            "FRK_SetRuntime".Work[#RootIndex].Payload.Info.RecordCount := #Slot;
        ELSIF #Phase = 2 THEN
            #Slot := "FRK_SetRecord"(RootIndex := #RootIndex, Scope := #Status.Name, WriteKey := "FRK_ConfigScratch".Entry.WriteKey);
            #Stored := "FRK_SetRuntime".Work[#RootIndex].Targets[#Slot];
            "FRK_ConfigCommit"(SlotIndex := #Stored, ModelCode := "FRK_SetRuntime".Work[#RootIndex].Payload.Info.ModelCode, Schema := "FRK_ConfigScratch".Schema, Record := "FRK_SetRuntime".Work[#RootIndex].Payload.Records[#Slot]);
        ELSE
            #Slot := "FRK_SetCheck"(RootIndex := #RootIndex, Scope := #Status.Name, Access := #Access, Ready := #Ready, WriteAccess := #Phase <> 3, ReserveTarget := #Phase = 1);
            IF #Slot = 0 THEN RETURN; END_IF;
            IF #Phase = 1 THEN
    #ConfigStageStationCfg.RequireTwoHandStart := "FRK_ConfigScratch".Value.Flag;
            END_IF;
        END_IF;
    END_IF;
    IF "FRK_SetRuntime".Work[#RootIndex].Payload.Info.Kind = 0 THEN
        "FRK_CfgDef_PressDemoUnit"(FieldIndex := 3);
        "FRK_SetRuntime".Work[#RootIndex].RejectScope := #Status.Name;
        "FRK_SetRuntime".Work[#RootIndex].RejectKey := "FRK_ConfigScratch".Entry.WriteKey;
        IF #Phase = 0 OR #Phase = 5 THEN
            IF #Phase = 5 AND NOT "FRK_ConfigDataAllowed"(Access := #Access, ForWrite := FALSE, Scope := #Status.Name) THEN RETURN; END_IF;
            IF #Phase = 5 AND (0 <> 0 OR "FRK_SetRuntime".Work[#RootIndex].Payload.Info.ModelCode = "FRK_ConfigStore".ActiveModels[#RootIndex]) THEN
    "FRK_ConfigScratch".Entry.ValueText := UDINT_TO_WSTRING(#ParCfg.IdealCycleMs);
                #Ok := "FRK_ConfigValidate"(Text := "FRK_ConfigScratch".Entry.ValueText);
            ELSE
                #Ok := "FRK_ConfigGet"(Scope := #Status.Name, ModelCode := "FRK_SetRuntime".Work[#RootIndex].Payload.Info.ModelCode);
            END_IF;
            IF NOT #Ok OR "FRK_SetRuntime".Work[#RootIndex].Payload.Info.RecordCount >= 21 THEN RETURN; END_IF;
            #Slot := "FRK_SetRuntime".Work[#RootIndex].Payload.Info.RecordCount + 1;
            "FRK_SetRuntime".Work[#RootIndex].Payload.Records[#Slot].Scope := #Status.Name;
            "FRK_SetRuntime".Work[#RootIndex].Payload.Records[#Slot].WriteKey := "FRK_ConfigScratch".Entry.WriteKey;
            "FRK_SetRuntime".Work[#RootIndex].Payload.Records[#Slot].Revision := "FRK_ConfigScratch".Entry.WriteRevision;
            "FRK_SetRuntime".Work[#RootIndex].Payload.Records[#Slot].Kind := "FRK_ConfigScratch".Entry.ConfigKind;
            "FRK_SetRuntime".Work[#RootIndex].Payload.Records[#Slot].ValueType := "FRK_ConfigScratch".Entry.ValueType;
            "FRK_SetRuntime".Work[#RootIndex].Payload.Records[#Slot].ValueText := WSTRING_TO_STRING("FRK_ConfigScratch".Entry.ValueText);
            "FRK_SetRuntime".Work[#RootIndex].Payload.Info.RecordCount := #Slot;
        ELSIF #Phase = 2 THEN
            #Slot := "FRK_SetRecord"(RootIndex := #RootIndex, Scope := #Status.Name, WriteKey := "FRK_ConfigScratch".Entry.WriteKey);
            #Stored := "FRK_SetRuntime".Work[#RootIndex].Targets[#Slot];
            "FRK_ConfigCommit"(SlotIndex := #Stored, ModelCode := "FRK_SetRuntime".Work[#RootIndex].Payload.Info.ModelCode, Schema := "FRK_ConfigScratch".Schema, Record := "FRK_SetRuntime".Work[#RootIndex].Payload.Records[#Slot]);
        ELSE
            #Slot := "FRK_SetCheck"(RootIndex := #RootIndex, Scope := #Status.Name, Access := #Access, Ready := #Ready, WriteAccess := #Phase <> 3, ReserveTarget := #Phase = 1);
            IF #Slot = 0 THEN RETURN; END_IF;
            IF #Phase = 1 THEN
    #ConfigStageParCfg.IdealCycleMs := LINT_TO_UDINT("FRK_ConfigScratch".Value.Number);
            END_IF;
        END_IF;
    END_IF;
    IF "FRK_SetRuntime".Work[#RootIndex].Payload.Info.Kind = 0 THEN
        "FRK_CfgDef_PressDemoUnit"(FieldIndex := 4);
        "FRK_SetRuntime".Work[#RootIndex].RejectScope := #Status.Name;
        "FRK_SetRuntime".Work[#RootIndex].RejectKey := "FRK_ConfigScratch".Entry.WriteKey;
        IF #Phase = 0 OR #Phase = 5 THEN
            IF #Phase = 5 AND NOT "FRK_ConfigDataAllowed"(Access := #Access, ForWrite := FALSE, Scope := #Status.Name) THEN RETURN; END_IF;
            IF #Phase = 5 AND (0 <> 0 OR "FRK_SetRuntime".Work[#RootIndex].Payload.Info.ModelCode = "FRK_ConfigStore".ActiveModels[#RootIndex]) THEN
    "FRK_ConfigScratch".Entry.ValueText := UDINT_TO_WSTRING(#ParCfg.BaselineWorkMs);
                #Ok := "FRK_ConfigValidate"(Text := "FRK_ConfigScratch".Entry.ValueText);
            ELSE
                #Ok := "FRK_ConfigGet"(Scope := #Status.Name, ModelCode := "FRK_SetRuntime".Work[#RootIndex].Payload.Info.ModelCode);
            END_IF;
            IF NOT #Ok OR "FRK_SetRuntime".Work[#RootIndex].Payload.Info.RecordCount >= 21 THEN RETURN; END_IF;
            #Slot := "FRK_SetRuntime".Work[#RootIndex].Payload.Info.RecordCount + 1;
            "FRK_SetRuntime".Work[#RootIndex].Payload.Records[#Slot].Scope := #Status.Name;
            "FRK_SetRuntime".Work[#RootIndex].Payload.Records[#Slot].WriteKey := "FRK_ConfigScratch".Entry.WriteKey;
            "FRK_SetRuntime".Work[#RootIndex].Payload.Records[#Slot].Revision := "FRK_ConfigScratch".Entry.WriteRevision;
            "FRK_SetRuntime".Work[#RootIndex].Payload.Records[#Slot].Kind := "FRK_ConfigScratch".Entry.ConfigKind;
            "FRK_SetRuntime".Work[#RootIndex].Payload.Records[#Slot].ValueType := "FRK_ConfigScratch".Entry.ValueType;
            "FRK_SetRuntime".Work[#RootIndex].Payload.Records[#Slot].ValueText := WSTRING_TO_STRING("FRK_ConfigScratch".Entry.ValueText);
            "FRK_SetRuntime".Work[#RootIndex].Payload.Info.RecordCount := #Slot;
        ELSIF #Phase = 2 THEN
            #Slot := "FRK_SetRecord"(RootIndex := #RootIndex, Scope := #Status.Name, WriteKey := "FRK_ConfigScratch".Entry.WriteKey);
            #Stored := "FRK_SetRuntime".Work[#RootIndex].Targets[#Slot];
            "FRK_ConfigCommit"(SlotIndex := #Stored, ModelCode := "FRK_SetRuntime".Work[#RootIndex].Payload.Info.ModelCode, Schema := "FRK_ConfigScratch".Schema, Record := "FRK_SetRuntime".Work[#RootIndex].Payload.Records[#Slot]);
        ELSE
            #Slot := "FRK_SetCheck"(RootIndex := #RootIndex, Scope := #Status.Name, Access := #Access, Ready := #Ready, WriteAccess := #Phase <> 3, ReserveTarget := #Phase = 1);
            IF #Slot = 0 THEN RETURN; END_IF;
            IF #Phase = 1 THEN
    #ConfigStageParCfg.BaselineWorkMs := LINT_TO_UDINT("FRK_ConfigScratch".Value.Number);
            END_IF;
        END_IF;
    END_IF;
    IF "FRK_SetRuntime".Work[#RootIndex].Payload.Info.Kind = 0 THEN
        "FRK_CfgDef_PressDemoUnit"(FieldIndex := 5);
        "FRK_SetRuntime".Work[#RootIndex].RejectScope := #Status.Name;
        "FRK_SetRuntime".Work[#RootIndex].RejectKey := "FRK_ConfigScratch".Entry.WriteKey;
        IF #Phase = 0 OR #Phase = 5 THEN
            IF #Phase = 5 AND NOT "FRK_ConfigDataAllowed"(Access := #Access, ForWrite := FALSE, Scope := #Status.Name) THEN RETURN; END_IF;
            IF #Phase = 5 AND (0 <> 0 OR "FRK_SetRuntime".Work[#RootIndex].Payload.Info.ModelCode = "FRK_ConfigStore".ActiveModels[#RootIndex]) THEN
    "FRK_ConfigScratch".Entry.ValueText := DINT_TO_WSTRING(TIME_TO_DINT(#ParCfg.Timeout));
                #Ok := "FRK_ConfigValidate"(Text := "FRK_ConfigScratch".Entry.ValueText);
            ELSE
                #Ok := "FRK_ConfigGet"(Scope := #Status.Name, ModelCode := "FRK_SetRuntime".Work[#RootIndex].Payload.Info.ModelCode);
            END_IF;
            IF NOT #Ok OR "FRK_SetRuntime".Work[#RootIndex].Payload.Info.RecordCount >= 21 THEN RETURN; END_IF;
            #Slot := "FRK_SetRuntime".Work[#RootIndex].Payload.Info.RecordCount + 1;
            "FRK_SetRuntime".Work[#RootIndex].Payload.Records[#Slot].Scope := #Status.Name;
            "FRK_SetRuntime".Work[#RootIndex].Payload.Records[#Slot].WriteKey := "FRK_ConfigScratch".Entry.WriteKey;
            "FRK_SetRuntime".Work[#RootIndex].Payload.Records[#Slot].Revision := "FRK_ConfigScratch".Entry.WriteRevision;
            "FRK_SetRuntime".Work[#RootIndex].Payload.Records[#Slot].Kind := "FRK_ConfigScratch".Entry.ConfigKind;
            "FRK_SetRuntime".Work[#RootIndex].Payload.Records[#Slot].ValueType := "FRK_ConfigScratch".Entry.ValueType;
            "FRK_SetRuntime".Work[#RootIndex].Payload.Records[#Slot].ValueText := WSTRING_TO_STRING("FRK_ConfigScratch".Entry.ValueText);
            "FRK_SetRuntime".Work[#RootIndex].Payload.Info.RecordCount := #Slot;
        ELSIF #Phase = 2 THEN
            #Slot := "FRK_SetRecord"(RootIndex := #RootIndex, Scope := #Status.Name, WriteKey := "FRK_ConfigScratch".Entry.WriteKey);
            #Stored := "FRK_SetRuntime".Work[#RootIndex].Targets[#Slot];
            "FRK_ConfigCommit"(SlotIndex := #Stored, ModelCode := "FRK_SetRuntime".Work[#RootIndex].Payload.Info.ModelCode, Schema := "FRK_ConfigScratch".Schema, Record := "FRK_SetRuntime".Work[#RootIndex].Payload.Records[#Slot]);
        ELSE
            #Slot := "FRK_SetCheck"(RootIndex := #RootIndex, Scope := #Status.Name, Access := #Access, Ready := #Ready, WriteAccess := #Phase <> 3, ReserveTarget := #Phase = 1);
            IF #Slot = 0 THEN RETURN; END_IF;
            IF #Phase = 1 THEN
    #ConfigStageParCfg.Timeout := DINT_TO_TIME(LINT_TO_DINT("FRK_ConfigScratch".Value.Number));
            END_IF;
        END_IF;
    END_IF;
    IF "FRK_SetRuntime".Work[#RootIndex].Payload.Info.Kind = 0 THEN
        "FRK_CfgDef_PressDemoUnit"(FieldIndex := 6);
        "FRK_SetRuntime".Work[#RootIndex].RejectScope := #Status.Name;
        "FRK_SetRuntime".Work[#RootIndex].RejectKey := "FRK_ConfigScratch".Entry.WriteKey;
        IF #Phase = 0 OR #Phase = 5 THEN
            IF #Phase = 5 AND NOT "FRK_ConfigDataAllowed"(Access := #Access, ForWrite := FALSE, Scope := #Status.Name) THEN RETURN; END_IF;
            IF #Phase = 5 AND (0 <> 0 OR "FRK_SetRuntime".Work[#RootIndex].Payload.Info.ModelCode = "FRK_ConfigStore".ActiveModels[#RootIndex]) THEN
    "FRK_ConfigScratch".Entry.ValueText := DINT_TO_WSTRING(TIME_TO_DINT(#ParCfg.TransferSettleTime));
                #Ok := "FRK_ConfigValidate"(Text := "FRK_ConfigScratch".Entry.ValueText);
            ELSE
                #Ok := "FRK_ConfigGet"(Scope := #Status.Name, ModelCode := "FRK_SetRuntime".Work[#RootIndex].Payload.Info.ModelCode);
            END_IF;
            IF NOT #Ok OR "FRK_SetRuntime".Work[#RootIndex].Payload.Info.RecordCount >= 21 THEN RETURN; END_IF;
            #Slot := "FRK_SetRuntime".Work[#RootIndex].Payload.Info.RecordCount + 1;
            "FRK_SetRuntime".Work[#RootIndex].Payload.Records[#Slot].Scope := #Status.Name;
            "FRK_SetRuntime".Work[#RootIndex].Payload.Records[#Slot].WriteKey := "FRK_ConfigScratch".Entry.WriteKey;
            "FRK_SetRuntime".Work[#RootIndex].Payload.Records[#Slot].Revision := "FRK_ConfigScratch".Entry.WriteRevision;
            "FRK_SetRuntime".Work[#RootIndex].Payload.Records[#Slot].Kind := "FRK_ConfigScratch".Entry.ConfigKind;
            "FRK_SetRuntime".Work[#RootIndex].Payload.Records[#Slot].ValueType := "FRK_ConfigScratch".Entry.ValueType;
            "FRK_SetRuntime".Work[#RootIndex].Payload.Records[#Slot].ValueText := WSTRING_TO_STRING("FRK_ConfigScratch".Entry.ValueText);
            "FRK_SetRuntime".Work[#RootIndex].Payload.Info.RecordCount := #Slot;
        ELSIF #Phase = 2 THEN
            #Slot := "FRK_SetRecord"(RootIndex := #RootIndex, Scope := #Status.Name, WriteKey := "FRK_ConfigScratch".Entry.WriteKey);
            #Stored := "FRK_SetRuntime".Work[#RootIndex].Targets[#Slot];
            "FRK_ConfigCommit"(SlotIndex := #Stored, ModelCode := "FRK_SetRuntime".Work[#RootIndex].Payload.Info.ModelCode, Schema := "FRK_ConfigScratch".Schema, Record := "FRK_SetRuntime".Work[#RootIndex].Payload.Records[#Slot]);
        ELSE
            #Slot := "FRK_SetCheck"(RootIndex := #RootIndex, Scope := #Status.Name, Access := #Access, Ready := #Ready, WriteAccess := #Phase <> 3, ReserveTarget := #Phase = 1);
            IF #Slot = 0 THEN RETURN; END_IF;
            IF #Phase = 1 THEN
    #ConfigStageParCfg.TransferSettleTime := DINT_TO_TIME(LINT_TO_DINT("FRK_ConfigScratch".Value.Number));
            END_IF;
        END_IF;
    END_IF;
    IF "FRK_SetRuntime".Work[#RootIndex].Payload.Info.Kind = 0 THEN
        "FRK_CfgDef_PressDemoUnit"(FieldIndex := 7);
        "FRK_SetRuntime".Work[#RootIndex].RejectScope := #Status.Name;
        "FRK_SetRuntime".Work[#RootIndex].RejectKey := "FRK_ConfigScratch".Entry.WriteKey;
        IF #Phase = 0 OR #Phase = 5 THEN
            IF #Phase = 5 AND NOT "FRK_ConfigDataAllowed"(Access := #Access, ForWrite := FALSE, Scope := #Status.Name) THEN RETURN; END_IF;
            IF #Phase = 5 AND (0 <> 0 OR "FRK_SetRuntime".Work[#RootIndex].Payload.Info.ModelCode = "FRK_ConfigStore".ActiveModels[#RootIndex]) THEN
    "FRK_ConfigScratch".Entry.ValueText := DINT_TO_WSTRING(TIME_TO_DINT(#ParCfg.PressSettleTime));
                #Ok := "FRK_ConfigValidate"(Text := "FRK_ConfigScratch".Entry.ValueText);
            ELSE
                #Ok := "FRK_ConfigGet"(Scope := #Status.Name, ModelCode := "FRK_SetRuntime".Work[#RootIndex].Payload.Info.ModelCode);
            END_IF;
            IF NOT #Ok OR "FRK_SetRuntime".Work[#RootIndex].Payload.Info.RecordCount >= 21 THEN RETURN; END_IF;
            #Slot := "FRK_SetRuntime".Work[#RootIndex].Payload.Info.RecordCount + 1;
            "FRK_SetRuntime".Work[#RootIndex].Payload.Records[#Slot].Scope := #Status.Name;
            "FRK_SetRuntime".Work[#RootIndex].Payload.Records[#Slot].WriteKey := "FRK_ConfigScratch".Entry.WriteKey;
            "FRK_SetRuntime".Work[#RootIndex].Payload.Records[#Slot].Revision := "FRK_ConfigScratch".Entry.WriteRevision;
            "FRK_SetRuntime".Work[#RootIndex].Payload.Records[#Slot].Kind := "FRK_ConfigScratch".Entry.ConfigKind;
            "FRK_SetRuntime".Work[#RootIndex].Payload.Records[#Slot].ValueType := "FRK_ConfigScratch".Entry.ValueType;
            "FRK_SetRuntime".Work[#RootIndex].Payload.Records[#Slot].ValueText := WSTRING_TO_STRING("FRK_ConfigScratch".Entry.ValueText);
            "FRK_SetRuntime".Work[#RootIndex].Payload.Info.RecordCount := #Slot;
        ELSIF #Phase = 2 THEN
            #Slot := "FRK_SetRecord"(RootIndex := #RootIndex, Scope := #Status.Name, WriteKey := "FRK_ConfigScratch".Entry.WriteKey);
            #Stored := "FRK_SetRuntime".Work[#RootIndex].Targets[#Slot];
            "FRK_ConfigCommit"(SlotIndex := #Stored, ModelCode := "FRK_SetRuntime".Work[#RootIndex].Payload.Info.ModelCode, Schema := "FRK_ConfigScratch".Schema, Record := "FRK_SetRuntime".Work[#RootIndex].Payload.Records[#Slot]);
        ELSE
            #Slot := "FRK_SetCheck"(RootIndex := #RootIndex, Scope := #Status.Name, Access := #Access, Ready := #Ready, WriteAccess := #Phase <> 3, ReserveTarget := #Phase = 1);
            IF #Slot = 0 THEN RETURN; END_IF;
            IF #Phase = 1 THEN
    #ConfigStageParCfg.PressSettleTime := DINT_TO_TIME(LINT_TO_DINT("FRK_ConfigScratch".Value.Number));
            END_IF;
        END_IF;
    END_IF;
    IF #Phase = 2 AND "FRK_SetRuntime".Work[#RootIndex].Payload.Info.Kind = 0 THEN #ParCfg := #ConfigStageParCfg; END_IF;
    IF #Phase = 2 AND "FRK_SetRuntime".Work[#RootIndex].Payload.Info.Kind = 1 THEN #StationCfg := #ConfigStageStationCfg; END_IF;
    #Ok := "FRK_CfgSetWalk_CylinderCM"(Module := #PressRam, RootIndex := #RootIndex, Phase := #Phase, Access := #Access, Ready := #Ready);
    IF NOT #Ok THEN RETURN; END_IF;
    #Ok := "FRK_CfgSetWalk_CylinderCM"(Module := #Door, RootIndex := #RootIndex, Phase := #Phase, Access := #Access, Ready := #Ready);
    IF NOT #Ok THEN RETURN; END_IF;
    #Ok := "FRK_CfgSetWalk_CylinderCM"(Module := #PartSlide, RootIndex := #RootIndex, Phase := #Phase, Access := #Access, Ready := #Ready);
    IF NOT #Ok THEN RETURN; END_IF;
    #Ok := "FRK_CfgSetWalk_TwoHandStartCM"(Module := #TwoHand, RootIndex := #RootIndex, Phase := #Phase, Access := #Access, Ready := #Ready);
    IF NOT #Ok THEN RETURN; END_IF;
    #Ok := "FRK_CfgSetWalk_DigitalInputCM"(Module := #PartPresentSensor, RootIndex := #RootIndex, Phase := #Phase, Access := #Access, Ready := #Ready);
    IF NOT #Ok THEN RETURN; END_IF;
    #Ok := "FRK_CfgSetWalk_AirPressureMonitorCM"(Module := #AirPressureMonitor, RootIndex := #RootIndex, Phase := #Phase, Access := #Access, Ready := #Ready);
    IF NOT #Ok THEN RETURN; END_IF;
    #FRK_CfgSetWalk_PressDemoUnit := TRUE;
END_FUNCTION
FUNCTION "FRK_CfgOperation_PressDemoUnit" : Void
{ S7_Optimized_Access := 'TRUE' }
VERSION : 0.1
VAR_IN_OUT
    Core : "FRK_Core";
    Status : "ST_ModuleStatus";
    ParCfg : "ST_PressDemoParCfg";
    ModePolicy : Array[0..6] of "ST_ModePolicy";
    Access : "FRK_Access";
    Unit : "FRK_Unit";
    HmiResponse : "ST_HmiResponse";
    AlarmLog : "FRK_AlarmLog";
    ConfigPersist : "ST_ConfigPersistStatus";
    ConfigCursor : "FRK_ConfigCursor";
    ConfigRev : UDInt;
    Model : "ST_ModelId";
    AvailableModelCount : Int;
    ConfigStaged : Bool;
    ModelCapacity : Int;
    SequenceStepDef : Array[1..23] of "ST_SequenceStepDef";
    SequenceStepCount : Int;
    SupportedModesPublished : Array[0..6] of Bool;
    StationCfg : "ST_PressDemoStationCfg";
    ConfigStageParCfg : "ST_PressDemoParCfg";
    ConfigDefaultParCfg : "ST_PressDemoParCfg";
    PressRam : "FB_CylinderCM";
    Door : "FB_CylinderCM";
    PartSlide : "FB_CylinderCM";
    TwoHand : "FB_TwoHandStartCM";
    PartPresentSensor : "FB_DigitalInputCM";
    AirPressureMonitor : "FB_AirPressureMonitorCM";
END_VAR
VAR_TEMP
    RootIndex : Int;
    Request : "ST_HmiRequest";
    Ready : Bool;
    Matched : Bool;
    Ok : Bool;
    Desired : String[64];
    Scope : String[80];
    Key : String[160];
END_VAR
BEGIN
    #RootIndex := "FRK_ConfigRoot"(RegIndex := #Core.RegIndex);
    IF #Core.ParentIndex <> 0 OR #RootIndex = 0 THEN RETURN; END_IF;
    #Model.ModelCode := "FRK_ConfigStore".ActiveModels[#RootIndex];
    IF NOT #Unit.RequestPending THEN RETURN; END_IF;
    #Request := #Unit.Request;
    #Ready := #Core.Exec = 0 AND NOT #Unit.ModePending AND NOT #Unit.Clearing AND "FRK_DescendantsReady"(OwnerIndex := #Core.RegIndex);
    CASE #Request.Kind OF
        23:
            "FRK_ConfigBegin"(Cursor := #ConfigCursor, Page := #HmiResponse.ConfigPage, PageIndex := #Request.IntValue, Revision := #ConfigRev);
            #HmiResponse.Accepted := FALSE;
            #HmiResponse.Diagnostic := WSTRING#'std.error.modelNotAvailable';
            IF #Request.DurationMs <= INT_TO_UDINT(#AvailableModelCount) AND #Request.IntValue >= 0 AND #Request.IntValue <= 32767 THEN
                "FRK_Config_PressDemoUnit"(Core := #Core, Status := #Status, ParCfg := #ParCfg, ModePolicy := #ModePolicy, AvailableModelCount := #AvailableModelCount, ModelCapacity := #ModelCapacity, SequenceStepDef := #SequenceStepDef, SequenceStepCount := #SequenceStepCount, StationCfg := #StationCfg, PressRam := #PressRam, Door := #Door, PartSlide := #PartSlide, TwoHand := #TwoHand, PartPresentSensor := #PartPresentSensor, AirPressureMonitor := #AirPressureMonitor, Access := #Access, RootIndex := #RootIndex, ModelIndex := #Request.DurationMs, Cursor := #ConfigCursor, Page := #HmiResponse.ConfigPage);
                "FRK_ConfigFinish"(Cursor := #ConfigCursor, Page := #HmiResponse.ConfigPage);
                #HmiResponse.Accepted := TRUE; #HmiResponse.Diagnostic := WSTRING#'';
            END_IF;
        19, 27:
            #HmiResponse.Accepted := FALSE;
            "FRK_ConfigScratch".RejectDescription := WSTRING#'std.error.recipeSchemaInvalid';
            "FRK_ConfigScratch".RejectReason := 2004;
            "FRK_ConfigScratch".CommittedScope := #Status.Name;
            #HmiResponse.Diagnostic := "FRK_ConfigScratch".RejectDescription;
            #ConfigPersist.LastRejectScope := #Status.Name;
            #ConfigPersist.LastRejectKey := #Request.NameValue;
            #HmiResponse.Report.Count := 0; #HmiResponse.Report.Released := TRUE;
            IF #Request.Kind = 27 THEN
                "FRK_ManualCommon"(Core := #Core, Unit := #Unit, Status := #Status, Report := #HmiResponse.Report);
                #Ready := #Ready AND #HmiResponse.Report.Released AND #Request.DurationMs = 0;
                IF NOT #Ready THEN
                    #HmiResponse.Diagnostic := WSTRING#'std.release.unitNotReady';
                    IF #HmiResponse.Report.Count = 0 THEN "FRK_ReleaseReason"(Report := #HmiResponse.Report, Description := #HmiResponse.Diagnostic, Reason := 2002, Path := STRING_TO_WSTRING(#Status.Name), Kind := 4); END_IF;
                    RETURN; END_IF;
            END_IF;
            IF #Request.DurationMs <= INT_TO_UDINT(#AvailableModelCount) THEN
                #Matched := FALSE;
                #HmiResponse.Accepted := "FRK_CfgWrite_PressDemoUnit"(Core := #Core, Status := #Status, ParCfg := #ParCfg, StationCfg := #StationCfg, PressRam := #PressRam, Door := #Door, PartSlide := #PartSlide, TwoHand := #TwoHand, PartPresentSensor := #PartPresentSensor, AirPressureMonitor := #AirPressureMonitor, Access := #Access, Request := #Request, RootIndex := #RootIndex, RootReady := #Ready, Matched := #Matched);
            END_IF;
            IF #HmiResponse.Accepted THEN
                "FRK_ConfigWriteAudit"(Scope := "FRK_ConfigScratch".CommittedScope, Key := #Request.NameValue, Value := "FRK_ConfigScratch".CommittedText, Captured := #Request.Kind = 27, User := #Unit.RequestUser, AlarmLog := #AlarmLog);
                #ConfigRev := "FRK_ConfigRevision"(Previous := #ConfigRev);
                #HmiResponse.Diagnostic := WSTRING#'';
                #ConfigPersist.LastRejectScope := ''; #ConfigPersist.LastRejectKey := '';
            ELSE
                #ConfigPersist.LastRejectScope := "FRK_ConfigScratch".CommittedScope;
                #HmiResponse.Diagnostic := "FRK_ConfigScratch".RejectDescription;
                "FRK_ReleaseReason"(Report := #HmiResponse.Report, Description := #HmiResponse.Diagnostic, Reason := "FRK_ConfigScratch".RejectReason, Path := STRING_TO_WSTRING("FRK_ConfigScratch".CommittedScope), Kind := 4);
            END_IF;
        4:
            #HmiResponse.Accepted := FALSE;
            #HmiResponse.Diagnostic := WSTRING#'std.error.modelNotAvailable';
            #Desired := '';
            #Desired := WSTRING_TO_STRING(#Request.TextValue);
            IF STRING_TO_WSTRING(#Desired) <> #Request.TextValue OR NOT "FRK_ModelKnown"(RootIndex := #RootIndex, Code := #Desired) THEN #Desired := ''; END_IF;
            "FRK_UnitRelease"(Core := #Core, Unit := #Unit, Status := #Status, Policy := #ModePolicy, Access := #Access, Supported := #SupportedModesPublished, Report := #HmiResponse.Report, Gate := 3, Desired := -1, Trusted := FALSE);
            IF #Desired <> '' AND #HmiResponse.Report.Released THEN
                #Scope := ''; #Key := '';
                #Ok := "FRK_CfgRecipe_PressDemoUnit"(Status := #Status, ParCfg := #ParCfg, ConfigStaged := #ConfigStaged, ConfigStageParCfg := #ConfigStageParCfg, ConfigDefaultParCfg := #ConfigDefaultParCfg, PressRam := #PressRam, Door := #Door, PartSlide := #PartSlide, TwoHand := #TwoHand, PartPresentSensor := #PartPresentSensor, AirPressureMonitor := #AirPressureMonitor, ModelCode := #Desired, Phase := 1, RejectScope := #Scope, RejectKey := #Key);
                IF #Ok THEN
                    #Ok := "FRK_CfgRecipe_PressDemoUnit"(Status := #Status, ParCfg := #ParCfg, ConfigStaged := #ConfigStaged, ConfigStageParCfg := #ConfigStageParCfg, ConfigDefaultParCfg := #ConfigDefaultParCfg, PressRam := #PressRam, Door := #Door, PartSlide := #PartSlide, TwoHand := #TwoHand, PartPresentSensor := #PartPresentSensor, AirPressureMonitor := #AirPressureMonitor, ModelCode := #Desired, Phase := 2, RejectScope := #Scope, RejectKey := #Key);
                    "FRK_ConfigSetActiveModel"(RootIndex := #RootIndex, ModelCode := #Desired);
                    #Model.ModelCode := #Desired;
                    #ConfigRev := "FRK_ConfigRevision"(Previous := #ConfigRev);
                    #HmiResponse.Accepted := TRUE; #HmiResponse.Diagnostic := WSTRING#'';
                ELSE
                    #ConfigPersist.LastRejectScope := #Scope; #ConfigPersist.LastRejectKey := #Key;
                    #Ok := "FRK_CfgRecipe_PressDemoUnit"(Status := #Status, ParCfg := #ParCfg, ConfigStaged := #ConfigStaged, ConfigStageParCfg := #ConfigStageParCfg, ConfigDefaultParCfg := #ConfigDefaultParCfg, PressRam := #PressRam, Door := #Door, PartSlide := #PartSlide, TwoHand := #TwoHand, PartPresentSensor := #PartPresentSensor, AirPressureMonitor := #AirPressureMonitor, ModelCode := #Desired, Phase := 0, RejectScope := #Scope, RejectKey := #Key);
                    #HmiResponse.Diagnostic := WSTRING#'std.error.recipeSchemaInvalid';
                    "FRK_Fault"(Core := #Core, Status := #Status, ReasonCode := 2004, Description := #HmiResponse.Diagnostic);
                    #Status.Diagnostic.SourcePath := STRING_TO_WSTRING(#Scope);
                END_IF;
            END_IF;
        31:
            #HmiResponse.Accepted := #Access.CurrentLevel >= 3;
            IF #HmiResponse.Accepted THEN "FRK_ConfigStore".Acknowledged[#RootIndex] := TRUE; "FRK_PersistAckRoot"(RootIndex := #RootIndex);
            ELSE #HmiResponse.Diagnostic := WSTRING#'std.error.configRestoreAckRefused'; END_IF;
        ELSE RETURN;
    END_CASE;
END_FUNCTION
FUNCTION "FRK_CfgSetOperation_PressDemoUnit" : Void
{ S7_Optimized_Access := 'TRUE' }
VERSION : 0.1
VAR_INPUT
    Startup : Bool;
END_VAR
VAR_IN_OUT
    Core : "FRK_Core";
    Status : "ST_ModuleStatus";
    ParCfg : "ST_PressDemoParCfg";
    ModePolicy : Array[0..6] of "ST_ModePolicy";
    Access : "FRK_Access";
    Unit : "FRK_Unit";
    HmiResponse : "ST_HmiResponse";
    ConfigPersist : "ST_ConfigPersistStatus";
    ConfigRev : UDInt;
    Model : "ST_ModelId";
    AvailableModelCount : Int;
    ConfigSets : Array[1..4] of "ST_ConfigSetInfo";
    ConfigSetCount : Int;
    ConfigSetDocument : WString;
    ConfigSetDocumentLine : Int;
    ConfigSetDocumentLines : Int;
    SupportedModesPublished : Array[0..6] of Bool;
    StationCfg : "ST_PressDemoStationCfg";
    ConfigStageParCfg : "ST_PressDemoParCfg";
    ConfigStageStationCfg : "ST_PressDemoStationCfg";
    PressRam : "FB_CylinderCM";
    Door : "FB_CylinderCM";
    PartSlide : "FB_CylinderCM";
    TwoHand : "FB_TwoHandStartCM";
    PartPresentSensor : "FB_DigitalInputCM";
    AirPressureMonitor : "FB_AirPressureMonitorCM";
END_VAR
VAR_TEMP
    RootIndex : Int;
    Request : "ST_HmiRequest";
    Ready : Bool;
    SetName : String[80];
    Slot : Int;
    Ok : Bool;
    Exporting : Bool;
    Stamp : DTL;
    ResultCode : Int;
END_VAR
BEGIN
    #RootIndex := "FRK_ConfigRoot"(RegIndex := #Core.RegIndex);
    IF #Core.ParentIndex <> 0 OR #RootIndex = 0 THEN RETURN; END_IF;
    IF #Startup THEN
        "FRK_SetRuntime".Work[#RootIndex].Importing := FALSE; "FRK_SetRuntime".Work[#RootIndex].Exporting := FALSE; "FRK_SetRuntime".Work[#RootIndex].Piece := WSTRING#'';
        IF "FRK_SetStore".SchemaVersion <> 1 THEN
            FOR #Slot := 1 TO 4 DO "FRK_SetStore".Sets[#RootIndex, #Slot].Info.Used := FALSE; END_FOR;
        END_IF;
    END_IF;
    IF "FRK_SetRuntime".Work[#RootIndex].Generation <> #Access.SessionGeneration THEN
        "FRK_SetRuntime".Work[#RootIndex].Importing := FALSE; "FRK_SetRuntime".Work[#RootIndex].Exporting := FALSE; "FRK_SetRuntime".Work[#RootIndex].Piece := WSTRING#'';
        "FRK_SetRuntime".Work[#RootIndex].Generation := #Access.SessionGeneration;
    END_IF;
    IF NOT #Unit.RequestPending THEN RETURN; END_IF;
    #Request := #Unit.Request;
    #Exporting := "FRK_SetRuntime".Work[#RootIndex].Exporting; "FRK_SetRuntime".Work[#RootIndex].Exporting := FALSE;
    IF #Request.Kind <> 33 THEN "FRK_SetRuntime".Work[#RootIndex].Importing := FALSE; "FRK_SetRuntime".Work[#RootIndex].Piece := WSTRING#''; END_IF;
    IF #Request.Kind <> 32 THEN "FRK_SetRuntime".Work[#RootIndex].Exporting := FALSE; END_IF;
    IF #Request.Kind <> 28 AND #Request.Kind <> 29 AND #Request.Kind <> 30 AND #Request.Kind <> 32 AND #Request.Kind <> 33 AND #Request.Kind <> 35 AND #Request.Kind <> 38 THEN RETURN; END_IF;
    #HmiResponse.Accepted := FALSE; #HmiResponse.Diagnostic := WSTRING#'std.error.configSetRejected';
    #ConfigPersist.LastRejectScope := #Status.Name; #ConfigPersist.LastRejectKey := '';
    "FRK_SetRuntime".Work[#RootIndex].RejectScope := #Status.Name; "FRK_SetRuntime".Work[#RootIndex].RejectKey := '';
    IF #Access.CurrentLevel < #Access.Policy.Required[11] THEN "FRK_SetRuntime".Work[#RootIndex].Importing := FALSE; "FRK_SetRuntime".Work[#RootIndex].Exporting := FALSE; "FRK_SetRuntime".Work[#RootIndex].Piece := WSTRING#''; RETURN; END_IF;
    IF "FRK_ConfigRuntime".Unavailable THEN "FRK_ConfigRuntime".Failed[#RootIndex] := TRUE; "FRK_SetRuntime".Work[#RootIndex].Importing := FALSE; "FRK_SetRuntime".Work[#RootIndex].Exporting := FALSE; "FRK_SetRuntime".Work[#RootIndex].Piece := WSTRING#''; RETURN; END_IF;
    #Ready := #Core.Exec = 0 AND NOT #Unit.ModePending AND NOT #Unit.Clearing AND "FRK_DescendantsReady"(OwnerIndex := #Core.RegIndex);
    #SetName := WSTRING_TO_STRING(#Request.TextValue);
    IF #Request.Kind <> 33 THEN
        IF LEN(#Request.TextValue) < 1 AND #Request.Kind <> 30 THEN RETURN; END_IF;
        IF LEN(#Request.TextValue) > 80 OR STRING_TO_WSTRING(#SetName) <> #Request.TextValue THEN RETURN; END_IF;
    END_IF;
    "FRK_SetRuntime".Work[#RootIndex].RejectScope := #Status.Name; "FRK_SetRuntime".Work[#RootIndex].RejectKey := '';
    CASE #Request.Kind OF
        30:
            #ConfigSetCount := 0;
            FOR #Slot := 1 TO 4 DO
                IF "FRK_SetStore".Sets[#RootIndex, #Slot].Info.Used THEN
                    #ConfigSetCount := #ConfigSetCount + 1;
                    #ConfigSets[#ConfigSetCount] := "FRK_SetStore".Sets[#RootIndex, #Slot].Info;
                END_IF;
            END_FOR;
            #HmiResponse.Accepted := TRUE;
        35:
            #Slot := "FRK_SetFind"(RootIndex := #RootIndex, SetName := #SetName);
            IF #Slot > 0 THEN "FRK_SetStore".Sets[#RootIndex, #Slot].Info.Used := FALSE; #HmiResponse.Accepted := TRUE; END_IF;
        28:
            #Slot := "FRK_SetSlot"(RootIndex := #RootIndex, SetName := #SetName);
            IF #Slot = 0 OR (#Request.IntValue <> 0 AND #Request.IntValue <> 1 AND #Request.IntValue <> 2) THEN RETURN; END_IF;
            "FRK_SetRuntime".Work[#RootIndex].Payload.Info.SetName := #SetName; "FRK_SetRuntime".Work[#RootIndex].Payload.Info.RootIdentity := #Status.Name;
            "FRK_SetRuntime".Work[#RootIndex].Payload.Info.SetSchema := 1; "FRK_SetRuntime".Work[#RootIndex].Payload.Info.ConfigRev := #ConfigRev;
            "FRK_SetRuntime".Work[#RootIndex].Payload.Info.Kind := #Request.IntValue; "FRK_SetRuntime".Work[#RootIndex].Payload.Info.RecordCount := 0;
            "FRK_SetRuntime".Work[#RootIndex].Payload.Info.ModelCode := '';
            IF #Request.IntValue = 0 THEN "FRK_SetRuntime".Work[#RootIndex].Payload.Info.ModelCode := #Model.ModelCode; END_IF;
            #ResultCode := RD_SYS_T(OUT => #Stamp); "FRK_SetRuntime".Work[#RootIndex].Payload.Info.CreatedAt := DTL_TO_LDT(#Stamp);
            "FRK_SetRuntime".Work[#RootIndex].Payload.Info.TimeSynchronized := FALSE; "FRK_SetRuntime".Work[#RootIndex].Payload.Info.Used := TRUE;
            #Ok := "FRK_CfgSetWalk_PressDemoUnit"(Status := #Status, ParCfg := #ParCfg, StationCfg := #StationCfg, ConfigStageParCfg := #ConfigStageParCfg, ConfigStageStationCfg := #ConfigStageStationCfg, PressRam := #PressRam, Door := #Door, PartSlide := #PartSlide, TwoHand := #TwoHand, PartPresentSensor := #PartPresentSensor, AirPressureMonitor := #AirPressureMonitor, RootIndex := #RootIndex, Phase := 0, Access := #Access, Ready := #Ready);
            IF #Ok THEN #Ok := "FRK_SetShape"(RootIndex := #RootIndex, RootIdentity := #Status.Name); END_IF;
            IF #Ok AND "FRK_SetRuntime".Work[#RootIndex].Payload.Info.RecordCount > 0 THEN "FRK_SetStore".Sets[#RootIndex, #Slot] := "FRK_SetRuntime".Work[#RootIndex].Payload; #HmiResponse.Accepted := TRUE; END_IF;
        29:
            #Slot := "FRK_SetFind"(RootIndex := #RootIndex, SetName := #SetName);
            IF #Slot = 0 THEN RETURN; END_IF;
            "FRK_SetRuntime".Work[#RootIndex].Payload := "FRK_SetStore".Sets[#RootIndex, #Slot];
            #Ok := "FRK_SetShape"(RootIndex := #RootIndex, RootIdentity := #Status.Name);
            IF NOT #Ok THEN RETURN; END_IF;
            IF "FRK_SetRuntime".Work[#RootIndex].Payload.Info.Kind = 0 THEN
                IF NOT "FRK_ModelKnown"(RootIndex := #RootIndex, Code := "FRK_SetRuntime".Work[#RootIndex].Payload.Info.ModelCode) THEN RETURN; END_IF;
                "FRK_UnitRelease"(Core := #Core, Unit := #Unit, Status := #Status, Policy := #ModePolicy, Access := #Access, Supported := #SupportedModesPublished, Report := #HmiResponse.Report, Gate := 3, Desired := -1, Trusted := FALSE);
                IF NOT #HmiResponse.Report.Released THEN RETURN; END_IF;
            END_IF;
            "FRK_SetValidateBegin"(RootIndex := #RootIndex); #Ok := "FRK_CfgSetWalk_PressDemoUnit"(Status := #Status, ParCfg := #ParCfg, StationCfg := #StationCfg, ConfigStageParCfg := #ConfigStageParCfg, ConfigStageStationCfg := #ConfigStageStationCfg, PressRam := #PressRam, Door := #Door, PartSlide := #PartSlide, TwoHand := #TwoHand, PartPresentSensor := #PartPresentSensor, AirPressureMonitor := #AirPressureMonitor, RootIndex := #RootIndex, Phase := 1, Access := #Access, Ready := #Ready);
            IF #Ok THEN #Ok := "FRK_SetValidateEnd"(RootIndex := #RootIndex); END_IF;
            IF #Ok AND "FRK_SetRuntime".Work[#RootIndex].Matched = "FRK_SetRuntime".Work[#RootIndex].Payload.Info.RecordCount THEN
                #Ok := "FRK_CfgSetWalk_PressDemoUnit"(Status := #Status, ParCfg := #ParCfg, StationCfg := #StationCfg, ConfigStageParCfg := #ConfigStageParCfg, ConfigStageStationCfg := #ConfigStageStationCfg, PressRam := #PressRam, Door := #Door, PartSlide := #PartSlide, TwoHand := #TwoHand, PartPresentSensor := #PartPresentSensor, AirPressureMonitor := #AirPressureMonitor, RootIndex := #RootIndex, Phase := 2, Access := #Access, Ready := #Ready);
                IF "FRK_SetRuntime".Work[#RootIndex].Payload.Info.Kind = 0 THEN "FRK_ConfigSetActiveModel"(RootIndex := #RootIndex, ModelCode := "FRK_SetRuntime".Work[#RootIndex].Payload.Info.ModelCode); #Model.ModelCode := "FRK_SetRuntime".Work[#RootIndex].Payload.Info.ModelCode; END_IF;
                #ConfigRev := "FRK_ConfigRevision"(Previous := #ConfigRev);
                #HmiResponse.Accepted := TRUE;
            END_IF;
        32:
            #ConfigSetDocument := WSTRING#''; #ConfigSetDocumentLine := -1; #ConfigSetDocumentLines := 0;
            IF #Request.IntValue < 0 THEN "FRK_SetRuntime".Work[#RootIndex].Exporting := FALSE; RETURN; END_IF;
            IF #Request.IntValue = 0 THEN
                IF #Request.NameValue <> '' THEN "FRK_SetRuntime".Work[#RootIndex].Exporting := FALSE; RETURN; END_IF;
                #Slot := "FRK_SetFind"(RootIndex := #RootIndex, SetName := #SetName); IF #Slot = 0 THEN RETURN; END_IF;
                "FRK_SetRuntime".Work[#RootIndex].Payload := "FRK_SetStore".Sets[#RootIndex, #Slot];
                "FRK_SetRuntime".Work[#RootIndex].CurrentExport := FALSE; "FRK_SetRuntime".Work[#RootIndex].ExportToken := '';
                "FRK_SetRuntime".Work[#RootIndex].NextLine := 0; #Exporting := TRUE;
            END_IF;
            IF ("FRK_SetRuntime".Work[#RootIndex].CurrentExport AND #Request.NameValue <> "FRK_SetRuntime".Work[#RootIndex].ExportToken) OR (NOT "FRK_SetRuntime".Work[#RootIndex].CurrentExport AND #Request.NameValue <> '') THEN "FRK_SetRuntime".Work[#RootIndex].Exporting := FALSE; RETURN; END_IF;
            IF NOT #Exporting OR #SetName <> "FRK_SetRuntime".Work[#RootIndex].Payload.Info.SetName OR #Request.IntValue <> "FRK_SetRuntime".Work[#RootIndex].NextLine OR #Request.IntValue > "FRK_SetRuntime".Work[#RootIndex].Payload.Info.RecordCount THEN RETURN; END_IF;
            #Ok := "FRK_SetShape"(RootIndex := #RootIndex, RootIdentity := #Status.Name);
            "FRK_SetValidateBegin"(RootIndex := #RootIndex);
            IF #Ok THEN #Ok := "FRK_CfgSetWalk_PressDemoUnit"(Status := #Status, ParCfg := #ParCfg, StationCfg := #StationCfg, ConfigStageParCfg := #ConfigStageParCfg, ConfigStageStationCfg := #ConfigStageStationCfg, PressRam := #PressRam, Door := #Door, PartSlide := #PartSlide, TwoHand := #TwoHand, PartPresentSensor := #PartPresentSensor, AirPressureMonitor := #AirPressureMonitor, RootIndex := #RootIndex, Phase := 3, Access := #Access, Ready := #Ready); END_IF;
            IF NOT #Ok OR "FRK_SetRuntime".Work[#RootIndex].Matched <> "FRK_SetRuntime".Work[#RootIndex].Payload.Info.RecordCount THEN "FRK_SetRuntime".Work[#RootIndex].Exporting := FALSE; RETURN; END_IF;
            IF #Request.IntValue = 0 THEN #Ok := "FRK_JsonHeader"(Data := "FRK_SetRuntime".Work[#RootIndex].Payload.Info, Line := #ConfigSetDocument);
            ELSE #Ok := "FRK_JsonRecord"(Data := "FRK_SetRuntime".Work[#RootIndex].Payload.Records[#Request.IntValue], Line := #ConfigSetDocument); END_IF;
            IF #Ok THEN #ConfigSetDocumentLine := DINT_TO_INT(#Request.IntValue); #ConfigSetDocumentLines := "FRK_SetRuntime".Work[#RootIndex].Payload.Info.RecordCount; "FRK_SetRuntime".Work[#RootIndex].NextLine := "FRK_SetRuntime".Work[#RootIndex].NextLine + 1; #HmiResponse.Accepted := TRUE; END_IF;
            "FRK_SetRuntime".Work[#RootIndex].Exporting := #Ok AND #Request.IntValue < "FRK_SetRuntime".Work[#RootIndex].Payload.Info.RecordCount;
        38:
            #ConfigSetDocument := WSTRING#''; #ConfigSetDocumentLine := -1; #ConfigSetDocumentLines := 0;
            IF NOT "FRK_ExportTokenValid"(Token := #Request.NameValue) OR (#Request.IntValue <> 0 AND #Request.IntValue <> 1 AND #Request.IntValue <> 2) THEN RETURN; END_IF;
            IF #Request.DurationMs > INT_TO_UDINT(#AvailableModelCount) OR (#Request.IntValue <> 0 AND #Request.DurationMs <> 0) THEN RETURN; END_IF;
            "FRK_SetRuntime".Work[#RootIndex].Payload.Info.SetName := #SetName; "FRK_SetRuntime".Work[#RootIndex].Payload.Info.RootIdentity := #Status.Name;
            "FRK_SetRuntime".Work[#RootIndex].Payload.Info.SetSchema := 1; "FRK_SetRuntime".Work[#RootIndex].Payload.Info.ConfigRev := #ConfigRev;
            "FRK_SetRuntime".Work[#RootIndex].Payload.Info.Kind := #Request.IntValue; "FRK_SetRuntime".Work[#RootIndex].Payload.Info.RecordCount := 0;
            "FRK_SetRuntime".Work[#RootIndex].Payload.Info.ModelCode := '';
            IF #Request.IntValue = 0 THEN "FRK_SetRuntime".Work[#RootIndex].Payload.Info.ModelCode := "FRK_ConfigModelCode"(RootIndex := #RootIndex, ModelIndex := #Request.DurationMs); END_IF;
            #ResultCode := RD_SYS_T(OUT => #Stamp); "FRK_SetRuntime".Work[#RootIndex].Payload.Info.CreatedAt := DTL_TO_LDT(#Stamp);
            "FRK_SetRuntime".Work[#RootIndex].Payload.Info.TimeSynchronized := FALSE; "FRK_SetRuntime".Work[#RootIndex].Payload.Info.Used := TRUE;
            #Ok := "FRK_CfgSetWalk_PressDemoUnit"(Status := #Status, ParCfg := #ParCfg, StationCfg := #StationCfg, ConfigStageParCfg := #ConfigStageParCfg, ConfigStageStationCfg := #ConfigStageStationCfg, PressRam := #PressRam, Door := #Door, PartSlide := #PartSlide, TwoHand := #TwoHand, PartPresentSensor := #PartPresentSensor, AirPressureMonitor := #AirPressureMonitor, RootIndex := #RootIndex, Phase := 5, Access := #Access, Ready := #Ready);
            IF #Ok THEN #Ok := "FRK_SetShape"(RootIndex := #RootIndex, RootIdentity := #Status.Name); END_IF;
            IF NOT #Ok OR "FRK_SetRuntime".Work[#RootIndex].Payload.Info.RecordCount = 0 THEN RETURN; END_IF;
            #Ok := "FRK_JsonHeader"(Data := "FRK_SetRuntime".Work[#RootIndex].Payload.Info, Line := #ConfigSetDocument);
            IF NOT #Ok THEN RETURN; END_IF;
            "FRK_SetRuntime".Work[#RootIndex].ExportToken := #Request.NameValue; "FRK_SetRuntime".Work[#RootIndex].CurrentExport := TRUE; "FRK_SetRuntime".Work[#RootIndex].NextLine := 1; "FRK_SetRuntime".Work[#RootIndex].Exporting := TRUE;
            #ConfigSetDocumentLine := 0; #ConfigSetDocumentLines := "FRK_SetRuntime".Work[#RootIndex].Payload.Info.RecordCount; #HmiResponse.Accepted := TRUE;
        33:
            #Ok := "FRK_SetImport"(RootIndex := #RootIndex, Request := #Request);
            IF #Ok AND #Request.BoolValue THEN
                #Ok := "FRK_SetShape"(RootIndex := #RootIndex, RootIdentity := #Status.Name);
                "FRK_SetValidateBegin"(RootIndex := #RootIndex);
                IF #Ok THEN #Ok := "FRK_CfgSetWalk_PressDemoUnit"(Status := #Status, ParCfg := #ParCfg, StationCfg := #StationCfg, ConfigStageParCfg := #ConfigStageParCfg, ConfigStageStationCfg := #ConfigStageStationCfg, PressRam := #PressRam, Door := #Door, PartSlide := #PartSlide, TwoHand := #TwoHand, PartPresentSensor := #PartPresentSensor, AirPressureMonitor := #AirPressureMonitor, RootIndex := #RootIndex, Phase := 4, Access := #Access, Ready := TRUE); END_IF;
                IF #Ok THEN #Ok := "FRK_SetValidateEnd"(RootIndex := #RootIndex); END_IF;
                #Slot := "FRK_SetSlot"(RootIndex := #RootIndex, SetName := "FRK_SetRuntime".Work[#RootIndex].Payload.Info.SetName);
                IF #Ok AND #Slot > 0 THEN "FRK_SetStore".Sets[#RootIndex, #Slot] := "FRK_SetRuntime".Work[#RootIndex].Payload; ELSE #Ok := FALSE; END_IF;
            END_IF;
            #HmiResponse.Accepted := #Ok;
            IF NOT #Ok THEN "FRK_SetRuntime".Work[#RootIndex].Importing := FALSE; "FRK_SetRuntime".Work[#RootIndex].Piece := WSTRING#''; END_IF;
        ELSE RETURN;
    END_CASE;
    IF #HmiResponse.Accepted THEN
        #HmiResponse.Diagnostic := WSTRING#''; "FRK_ConfigRuntime".Failed[#RootIndex] := FALSE;
        #ConfigPersist.LastSetName := "FRK_SetRuntime".Work[#RootIndex].Payload.Info.SetName; #ConfigPersist.LastSetRecords := "FRK_SetRuntime".Work[#RootIndex].Payload.Info.RecordCount;
        #ConfigPersist.LastRejectScope := ''; #ConfigPersist.LastRejectKey := '';
    ELSE #ConfigPersist.LastRejectScope := "FRK_SetRuntime".Work[#RootIndex].RejectScope; #ConfigPersist.LastRejectKey := "FRK_SetRuntime".Work[#RootIndex].RejectKey; END_IF;
    IF #HmiResponse.Accepted AND (#Request.Kind = 28 OR #Request.Kind = 35 OR (#Request.Kind = 33 AND #Request.BoolValue)) THEN
        "FRK_PersistSetDirty"(RootIndex := #RootIndex, Ordinal := #Slot);
    END_IF;
END_FUNCTION
FUNCTION "FRK_CfgModelOperation_PressDemoUnit" : Void
{ S7_Optimized_Access := 'TRUE' }
VERSION : 0.1
VAR_IN_OUT
    Core : "FRK_Core";
    Status : "ST_ModuleStatus";
    ParCfg : "ST_PressDemoParCfg";
    Access : "FRK_Access";
    Unit : "FRK_Unit";
    HmiResponse : "ST_HmiResponse";
    AlarmLog : "FRK_AlarmLog";
    ConfigPersist : "ST_ConfigPersistStatus";
    ConfigRev : UDInt;
    AvailableModelCount : Int;
    ModelCapacity : Int;
    ModelGenerationSeen : UDInt;
    AvailableModels : Array[1..4] of "ST_ModelId";
    StationCfg : "ST_PressDemoStationCfg";
    ConfigStageParCfg : "ST_PressDemoParCfg";
    ConfigStageStationCfg : "ST_PressDemoStationCfg";
    PressRam : "FB_CylinderCM";
    Door : "FB_CylinderCM";
    PartSlide : "FB_CylinderCM";
    TwoHand : "FB_TwoHandStartCM";
    PartPresentSensor : "FB_DigitalInputCM";
    AirPressureMonitor : "FB_AirPressureMonitorCM";
END_VAR
VAR_TEMP
    RootIndex : Int;
    Index : Int;
    Slot : Int;
    Request : "ST_HmiRequest";
    NewCode : String[64];
    SourceCode : String[64];
    SetName : String[80];
    Ok : Bool;
    NativeResult : Int;
END_VAR
BEGIN
    #RootIndex := "FRK_ConfigRoot"(RegIndex := #Core.RegIndex);
    IF #Core.ParentIndex <> 0 OR #RootIndex = 0 THEN RETURN; END_IF;
    IF "FRK_ModelTick"(RootIndex := #RootIndex) THEN #ConfigRev := "FRK_ConfigRevision"(Previous := #ConfigRev); END_IF;
    #ModelCapacity := 4;
    #AvailableModelCount := "FRK_ModelStore".Rows[#RootIndex].Count;
    IF #ModelGenerationSeen <> "FRK_ModelStore".Rows[#RootIndex].Generation THEN
        FOR #Index := 1 TO 4 DO #AvailableModels[#Index].ModelCode := "FRK_ModelStore".Rows[#RootIndex].Codes[#Index]; END_FOR;
        #ModelGenerationSeen := "FRK_ModelStore".Rows[#RootIndex].Generation;
    END_IF;
    IF NOT #Unit.RequestPending OR #Unit.Request.Kind <> 37 THEN RETURN; END_IF;
    #Request := #Unit.Request;
    #HmiResponse.Accepted := FALSE; #HmiResponse.Diagnostic := WSTRING#'std.error.configSetRejected';
    #HmiResponse.Report.Count := 0; #HmiResponse.Report.Released := TRUE;
    "FRK_ReleaseReason"(Report := #HmiResponse.Report, Description := #HmiResponse.Diagnostic, Reason := 2002, Path := STRING_TO_WSTRING(#Status.Name), Kind := 4);
    #ConfigPersist.LastRejectScope := #Status.Name; #ConfigPersist.LastRejectKey := '';
    "FRK_SetRuntime".Work[#RootIndex].Importing := FALSE; "FRK_SetRuntime".Work[#RootIndex].Exporting := FALSE; "FRK_SetRuntime".Work[#RootIndex].Piece := WSTRING#'';
    IF #Access.CurrentLevel < #Access.Policy.Required[11] THEN
        #HmiResponse.Diagnostic := WSTRING#'std.error.accessDenied';
        #HmiResponse.Report.Count := 0; #HmiResponse.Report.Released := TRUE;
        "FRK_ReleaseReason"(Report := #HmiResponse.Report, Description := #HmiResponse.Diagnostic, Reason := 2002, Path := STRING_TO_WSTRING(#Status.Name), Kind := 1);
        RETURN;
    END_IF;
    IF NOT "FRK_ModelRuntime".Rows[#RootIndex].Ready OR "FRK_ModelRuntime".Rows[#RootIndex].State <> 0 OR "FRK_ConfigRuntime".Unavailable
        OR ("FRK_ConfigStore".Lost[#RootIndex] AND NOT "FRK_ConfigStore".Acknowledged[#RootIndex])
        OR "FRK_ModelStore".Rows[#RootIndex].Count >= 4 THEN RETURN; END_IF;
    IF LEN(#Request.NameValue) > 64 THEN RETURN; END_IF;
    #NewCode := #Request.NameValue;
    IF NOT "FRK_ModelCodeValid"(Code := #NewCode) OR "FRK_ModelKnown"(RootIndex := #RootIndex, Code := #NewCode)
        OR #Request.DurationMs <> 0 OR #Request.TargetPath <> WSTRING#'' THEN RETURN; END_IF;
    IF #Request.BoolValue THEN
        #SetName := WSTRING_TO_STRING(#Request.TextValue);
        IF LEN(#Request.TextValue) < 1 OR LEN(#Request.TextValue) > 80 OR STRING_TO_WSTRING(#SetName) <> #Request.TextValue THEN RETURN; END_IF;
        #Slot := "FRK_SetFind"(RootIndex := #RootIndex, SetName := #SetName); IF #Slot = 0 THEN RETURN; END_IF;
        "FRK_SetRuntime".Work[#RootIndex].Payload := "FRK_SetStore".Sets[#RootIndex, #Slot];
    ELSE
        IF #Request.IntValue < 0 OR #Request.TextValue <> WSTRING#'' THEN RETURN; END_IF;
        #SourceCode := "FRK_ConfigModelCode"(RootIndex := #RootIndex, ModelIndex := DINT_TO_UDINT(#Request.IntValue));
        IF #SourceCode = '' THEN RETURN; END_IF;
        "FRK_SetRuntime".Work[#RootIndex].Payload.Info.Used := TRUE; "FRK_SetRuntime".Work[#RootIndex].Payload.Info.SetSchema := 1;
        "FRK_SetRuntime".Work[#RootIndex].Payload.Info.RootIdentity := #Status.Name; "FRK_SetRuntime".Work[#RootIndex].Payload.Info.SetName := 'clone';
        "FRK_SetRuntime".Work[#RootIndex].Payload.Info.ConfigRev := #ConfigRev; "FRK_SetRuntime".Work[#RootIndex].Payload.Info.Kind := 0;
        "FRK_SetRuntime".Work[#RootIndex].Payload.Info.ModelCode := #SourceCode; "FRK_SetRuntime".Work[#RootIndex].Payload.Info.RecordCount := 0;
        #Ok := "FRK_CfgSetWalk_PressDemoUnit"(Status := #Status, ParCfg := #ParCfg, StationCfg := #StationCfg, ConfigStageParCfg := #ConfigStageParCfg, ConfigStageStationCfg := #ConfigStageStationCfg, PressRam := #PressRam, Door := #Door, PartSlide := #PartSlide, TwoHand := #TwoHand, PartPresentSensor := #PartPresentSensor, AirPressureMonitor := #AirPressureMonitor, RootIndex := #RootIndex, Phase := 0, Access := #Access, Ready := TRUE); IF NOT #Ok THEN RETURN; END_IF;
    END_IF;
    IF "FRK_SetRuntime".Work[#RootIndex].Payload.Info.Kind <> 0 OR NOT "FRK_ModelCodeValid"(Code := "FRK_SetRuntime".Work[#RootIndex].Payload.Info.ModelCode) THEN RETURN; END_IF;
    #Ok := "FRK_SetShape"(RootIndex := #RootIndex, RootIdentity := #Status.Name);
    IF NOT #Ok THEN RETURN; END_IF;
    "FRK_SetValidateBegin"(RootIndex := #RootIndex); #Ok := "FRK_CfgSetWalk_PressDemoUnit"(Status := #Status, ParCfg := #ParCfg, StationCfg := #StationCfg, ConfigStageParCfg := #ConfigStageParCfg, ConfigStageStationCfg := #ConfigStageStationCfg, PressRam := #PressRam, Door := #Door, PartSlide := #PartSlide, TwoHand := #TwoHand, PartPresentSensor := #PartPresentSensor, AirPressureMonitor := #AirPressureMonitor, RootIndex := #RootIndex, Phase := 3, Access := #Access, Ready := TRUE);
    IF #Ok THEN #Ok := "FRK_SetValidateEnd"(RootIndex := #RootIndex); END_IF;
    IF #Ok THEN "FRK_SetValidateBegin"(RootIndex := #RootIndex); #Ok := "FRK_CfgSetWalk_PressDemoUnit"(Status := #Status, ParCfg := #ParCfg, StationCfg := #StationCfg, ConfigStageParCfg := #ConfigStageParCfg, ConfigStageStationCfg := #ConfigStageStationCfg, PressRam := #PressRam, Door := #Door, PartSlide := #PartSlide, TwoHand := #TwoHand, PartPresentSensor := #PartPresentSensor, AirPressureMonitor := #AirPressureMonitor, RootIndex := #RootIndex, Phase := 4, Access := #Access, Ready := TRUE); END_IF;
    IF #Ok THEN #Ok := "FRK_SetValidateEnd"(RootIndex := #RootIndex); END_IF;
    IF NOT #Ok THEN
        #ConfigPersist.LastRejectScope := "FRK_SetRuntime".Work[#RootIndex].RejectScope;
        #ConfigPersist.LastRejectKey := "FRK_SetRuntime".Work[#RootIndex].RejectKey; RETURN;
    END_IF;
    FOR #Index := 1 TO "FRK_SetRuntime".Work[#RootIndex].Payload.Info.RecordCount DO
        #Slot := "FRK_ConfigReserve"(Scope := "FRK_SetRuntime".Work[#RootIndex].Payload.Records[#Index].Scope, Key := "FRK_SetRuntime".Work[#RootIndex].Payload.Records[#Index].WriteKey, ModelCode := #NewCode, Reserved := "FRK_SetRuntime".Work[#RootIndex].Targets);
        IF #Slot < 1 OR #Slot > 22 THEN RETURN; END_IF;
        "FRK_SetRuntime".Work[#RootIndex].Targets[#Index] := #Slot;
    END_FOR;
    FOR #Index := 1 TO "FRK_SetRuntime".Work[#RootIndex].Payload.Info.RecordCount DO
        "FRK_ConfigCommit"(SlotIndex := "FRK_SetRuntime".Work[#RootIndex].Targets[#Index], ModelCode := #NewCode, Schema := "FRK_SetRuntime".Work[#RootIndex].Schemas[#Index], Record := "FRK_SetRuntime".Work[#RootIndex].Payload.Records[#Index]);
    END_FOR;
    "FRK_ModelRuntime".Rows[#RootIndex].Stage := "FRK_ModelStore".Rows[#RootIndex];
    "FRK_ModelRuntime".Rows[#RootIndex].Stage.Count := "FRK_ModelRuntime".Rows[#RootIndex].Stage.Count + 1;
    "FRK_ModelRuntime".Rows[#RootIndex].Stage.Codes["FRK_ModelRuntime".Rows[#RootIndex].Stage.Count] := #NewCode;
    "FRK_ModelRuntime".Rows[#RootIndex].Stage.Generation := "FRK_ConfigRevision"(Previous := "FRK_ModelRuntime".Rows[#RootIndex].Stage.Generation);
    "FRK_ModelRuntime".Rows[#RootIndex].Stage.Checksum := "FRK_ModelCrc"(Catalog := "FRK_ModelRuntime".Rows[#RootIndex].Stage);
    "FRK_ModelRuntime".Rows[#RootIndex].State := 1;
    #NativeResult := RD_SYS_T(OUT => "FRK_ModelRuntime".Rows[#RootIndex].PendingSince);
    "FRK_ModelSave"(RootIndex := #RootIndex);
    #HmiResponse.Accepted := TRUE; #HmiResponse.Diagnostic := WSTRING#'';
    #HmiResponse.Report.Count := 0; #HmiResponse.Report.Released := TRUE;
    #ConfigPersist.LastRejectScope := ''; #ConfigPersist.LastRejectKey := '';
    "FRK_ConfigWriteAudit"(Scope := #Status.Name, Key := 'ModelCreation', Value := STRING_TO_WSTRING(#NewCode), Captured := FALSE, User := #Unit.RequestUser, AlarmLog := #AlarmLog);
END_FUNCTION
